(* Schneider Machine Expert - Basic project m200-cpp EXPERIMENTAL, file version 3.0.0.0 *)
(* ProjectInformations: Name=New project *)

HARDWARE
  Cpu 0: TM200CE40T
  EthernetConfiguration: NetworkName=M200, IpAllocationMode=FixedAddress, IpAddress=0.0.0.0, SubnetMask=0.0.0.0
  SerialLineConfiguration: Baud=Baud19200, Parity=ParityEven, DataBits=DataBits8, StopBits=StopBits1, PhysicalMedium=PhysicalMediumRs485, TransmissionMode=TransmissionModeModbusRtu, SlaveId=1, Addressing=SlaveAddressing
  MastTask: UsePeriodScanMode=false, PeriodScan=100
  FastTask: Period=255
  CpuBehavior: StartingMode=StartAsPreviousState, AutoSaveRamOnEeprom=true, WatchdogPeriod=250

SYMBOLS  (address, symbol, comment, settings)
  %S13      SB_FIRSTRUN  "Indicates the first controller cycle in RUN mode"
  %R0         [Type=Fifo]
  %R1         [Type=Lifo]
  %M0       compiler_reused_M0_0

POU Generated C++ - EXPERIMENTAL
  (* SectionNumber=0 *)

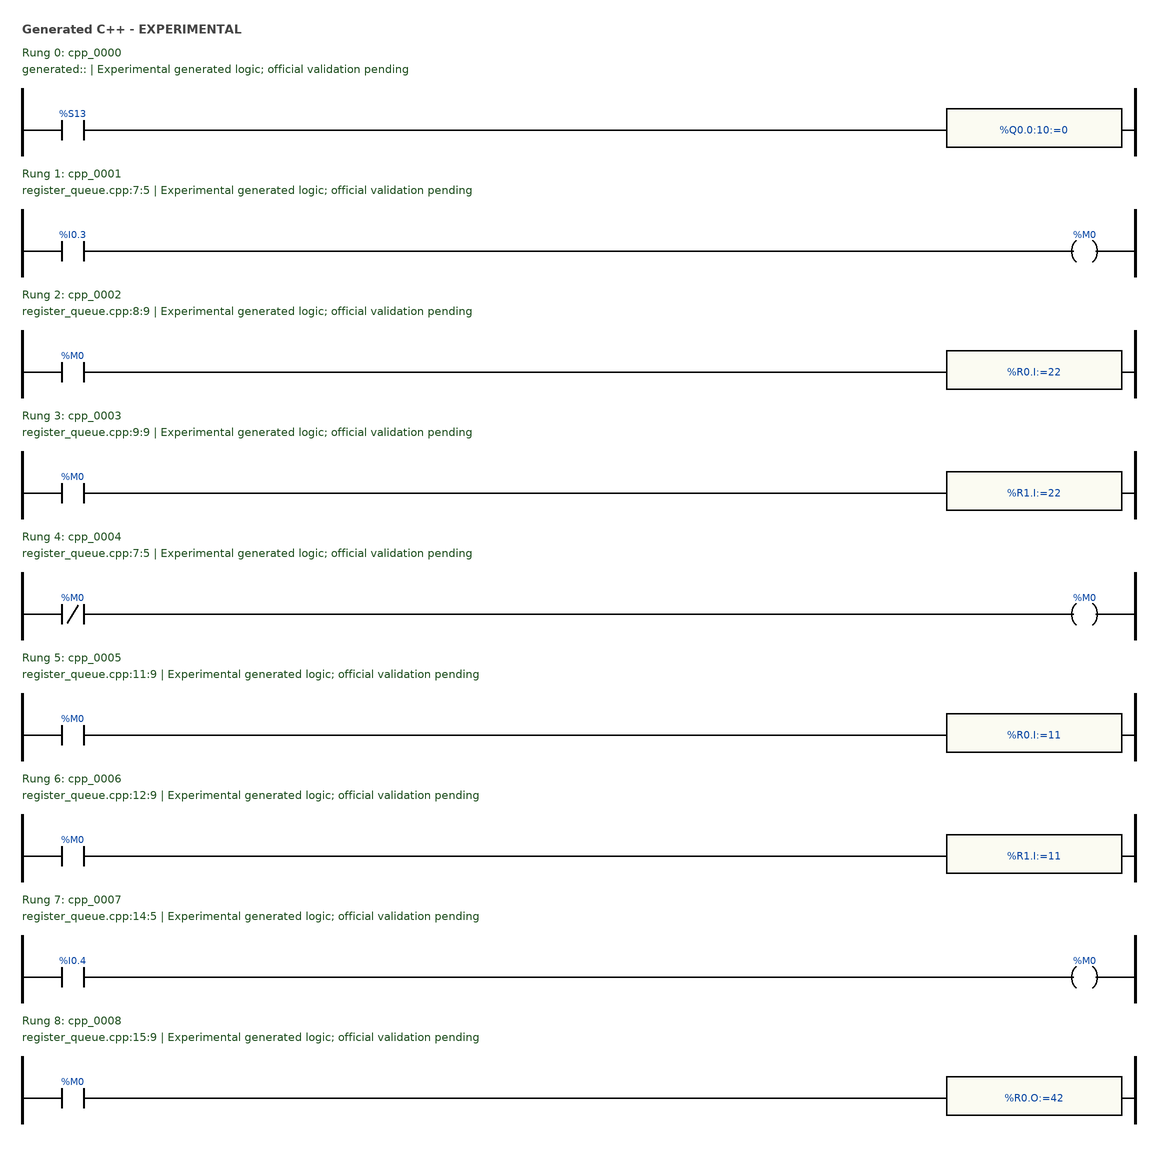

// Rung 0: cpp_0000
// generated:: | Experimental generated logic; official validation pending
  LD %S13                 (* SB_FIRSTRUN *)
  [%Q0.0:10:=0]
  // as ST:
  //   IF SB_FIRSTRUN THEN %Q0.0:10:=0; END_IF;

// Rung 1: cpp_0001
// register_queue.cpp:7:5 | Experimental generated logic; official validation pending
  LD %I0.3
  ST %M0                  (* compiler_reused_M0_0 *)
  // as ST:
  //   compiler_reused_M0_0 := %I0.3;

// Rung 2: cpp_0002
// register_queue.cpp:8:9 | Experimental generated logic; official validation pending
  LD %M0                  (* compiler_reused_M0_0 *)
  [%R0.I:=22]
  // as ST:
  //   IF compiler_reused_M0_0 THEN %R0.I:=22; END_IF;

// Rung 3: cpp_0003
// register_queue.cpp:9:9 | Experimental generated logic; official validation pending
  LD %M0                  (* compiler_reused_M0_0 *)
  [%R1.I:=22]
  // as ST:
  //   IF compiler_reused_M0_0 THEN %R1.I:=22; END_IF;

// Rung 4: cpp_0004
// register_queue.cpp:7:5 | Experimental generated logic; official validation pending
  LDN %M0                 (* compiler_reused_M0_0 *)
  ST %M0                  (* compiler_reused_M0_0 *)
  // as ST:
  //   compiler_reused_M0_0 := NOT compiler_reused_M0_0;

// Rung 5: cpp_0005
// register_queue.cpp:11:9 | Experimental generated logic; official validation pending
  LD %M0                  (* compiler_reused_M0_0 *)
  [%R0.I:=11]
  // as ST:
  //   IF compiler_reused_M0_0 THEN %R0.I:=11; END_IF;

// Rung 6: cpp_0006
// register_queue.cpp:12:9 | Experimental generated logic; official validation pending
  LD %M0                  (* compiler_reused_M0_0 *)
  [%R1.I:=11]
  // as ST:
  //   IF compiler_reused_M0_0 THEN %R1.I:=11; END_IF;

// Rung 7: cpp_0007
// register_queue.cpp:14:5 | Experimental generated logic; official validation pending
  LD %I0.4
  ST %M0                  (* compiler_reused_M0_0 *)
  // as ST:
  //   compiler_reused_M0_0 := %I0.4;

// Rung 8: cpp_0008
// register_queue.cpp:15:9 | Experimental generated logic; official validation pending
  LD %M0                  (* compiler_reused_M0_0 *)
  [%R0.O:=42]
  // as ST:
  //   IF compiler_reused_M0_0 THEN %R0.O:=42; END_IF;

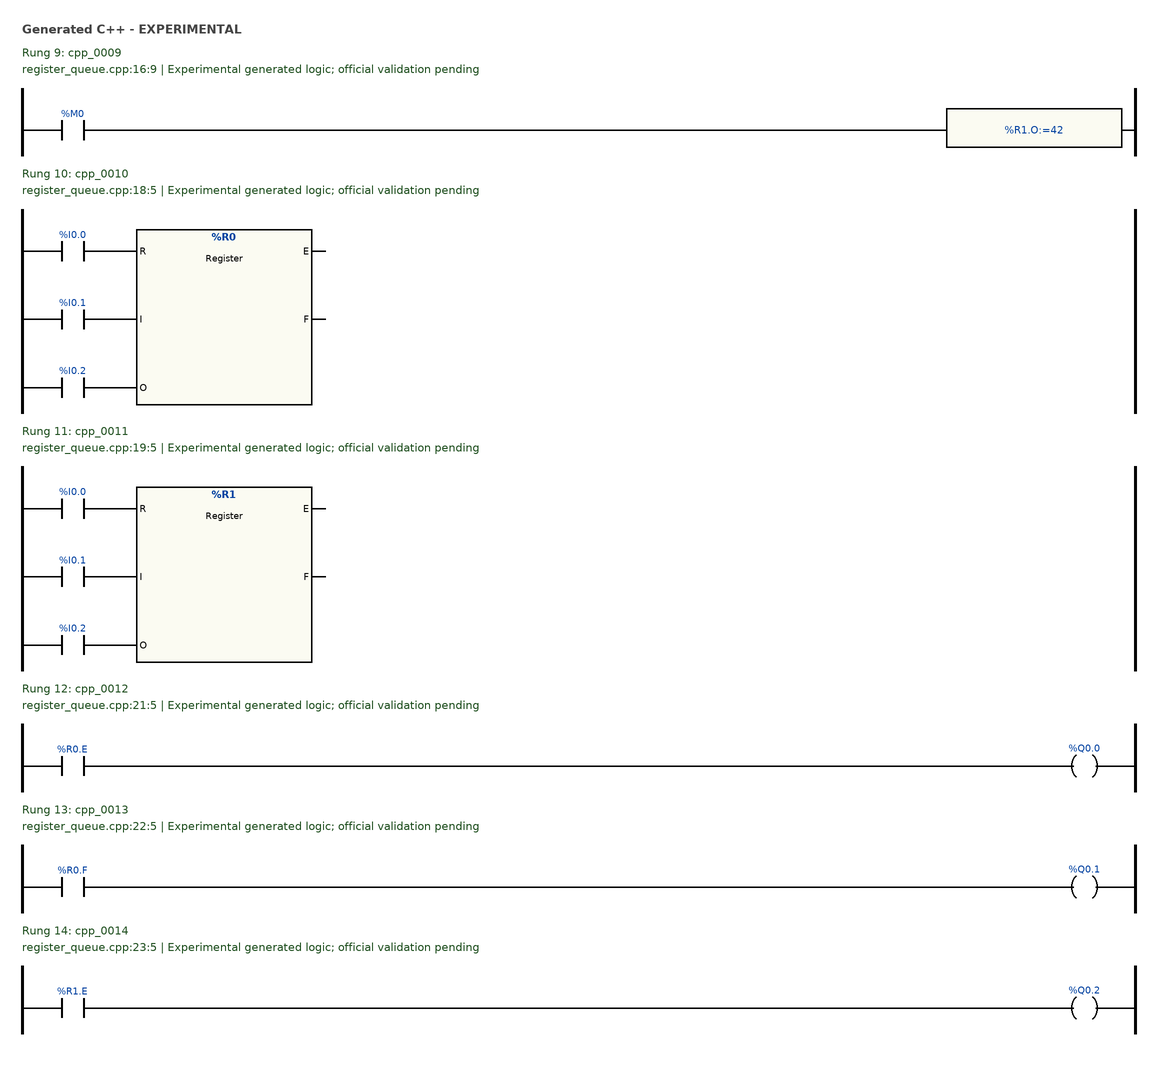

// Rung 9: cpp_0009
// register_queue.cpp:16:9 | Experimental generated logic; official validation pending
  LD %M0                  (* compiler_reused_M0_0 *)
  [%R1.O:=42]
  // as ST:
  //   IF compiler_reused_M0_0 THEN %R1.O:=42; END_IF;

// Rung 10: cpp_0010
// register_queue.cpp:18:5 | Experimental generated logic; official validation pending
  BLK %R0
  LD %I0.0
  R
  LD %I0.1
  I
  LD %I0.2
  O
  END_BLK
  // as ST:
  //   %R0(R := %I0.0, I := %I0.1, O := %I0.2);

// Rung 11: cpp_0011
// register_queue.cpp:19:5 | Experimental generated logic; official validation pending
  BLK %R1
  LD %I0.0
  R
  LD %I0.1
  I
  LD %I0.2
  O
  END_BLK
  // as ST:
  //   %R1(R := %I0.0, I := %I0.1, O := %I0.2);

// Rung 12: cpp_0012
// register_queue.cpp:21:5 | Experimental generated logic; official validation pending
  LD %R0.E
  ST %Q0.0
  // as ST:
  //   %Q0.0 := %R0.E;

// Rung 13: cpp_0013
// register_queue.cpp:22:5 | Experimental generated logic; official validation pending
  LD %R0.F
  ST %Q0.1
  // as ST:
  //   %Q0.1 := %R0.F;

// Rung 14: cpp_0014
// register_queue.cpp:23:5 | Experimental generated logic; official validation pending
  LD %R1.E
  ST %Q0.2
  // as ST:
  //   %Q0.2 := %R1.E;

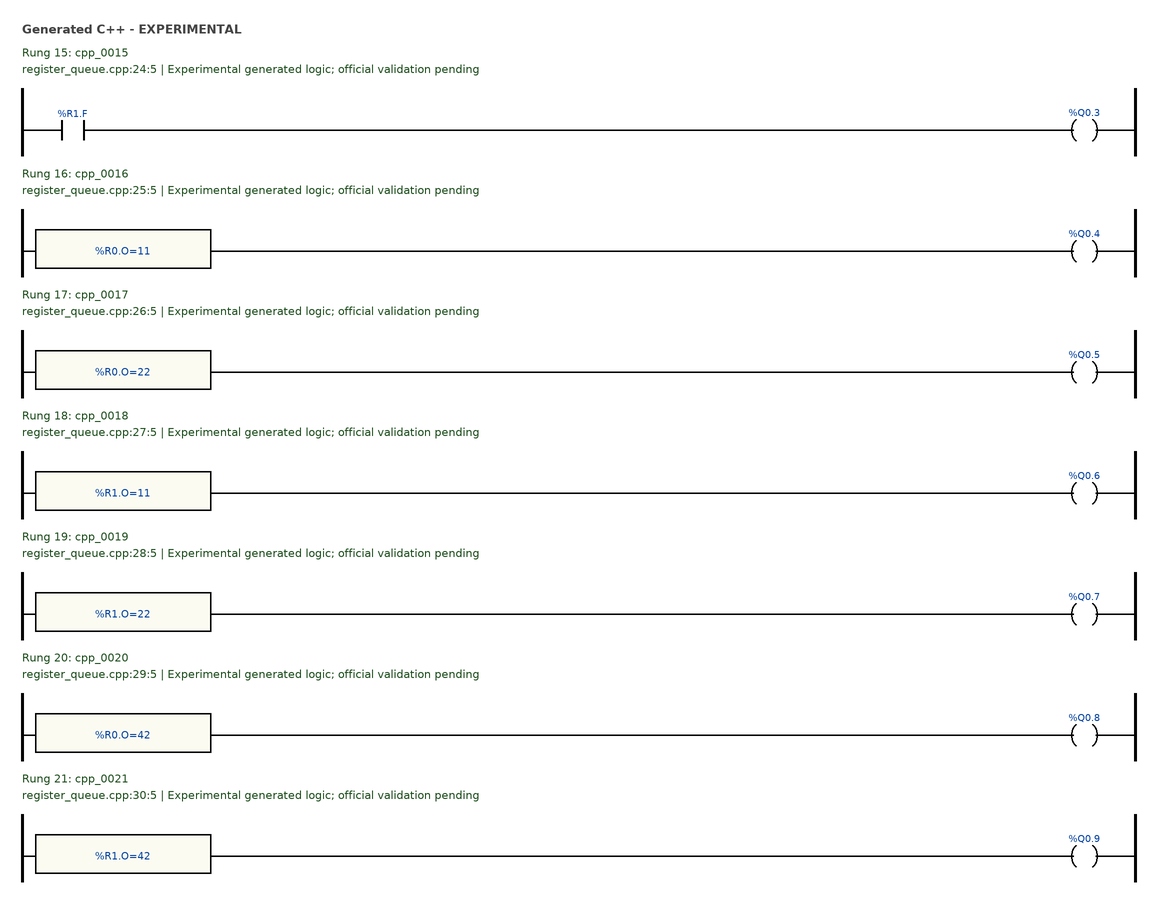

// Rung 15: cpp_0015
// register_queue.cpp:24:5 | Experimental generated logic; official validation pending
  LD %R1.F
  ST %Q0.3
  // as ST:
  //   %Q0.3 := %R1.F;

// Rung 16: cpp_0016
// register_queue.cpp:25:5 | Experimental generated logic; official validation pending
  LD [%R0.O=11]
  ST %Q0.4
  // as ST:
  //   %Q0.4 := %R0.O=11;

// Rung 17: cpp_0017
// register_queue.cpp:26:5 | Experimental generated logic; official validation pending
  LD [%R0.O=22]
  ST %Q0.5
  // as ST:
  //   %Q0.5 := %R0.O=22;

// Rung 18: cpp_0018
// register_queue.cpp:27:5 | Experimental generated logic; official validation pending
  LD [%R1.O=11]
  ST %Q0.6
  // as ST:
  //   %Q0.6 := %R1.O=11;

// Rung 19: cpp_0019
// register_queue.cpp:28:5 | Experimental generated logic; official validation pending
  LD [%R1.O=22]
  ST %Q0.7
  // as ST:
  //   %Q0.7 := %R1.O=22;

// Rung 20: cpp_0020
// register_queue.cpp:29:5 | Experimental generated logic; official validation pending
  LD [%R0.O=42]
  ST %Q0.8
  // as ST:
  //   %Q0.8 := %R0.O=42;

// Rung 21: cpp_0021
// register_queue.cpp:30:5 | Experimental generated logic; official validation pending
  LD [%R1.O=42]
  ST %Q0.9
  // as ST:
  //   %Q0.9 := %R1.O=42;
